Fanuc KAREL source: kd00006.KL

-- PROVISIONAL review KL for V770-1; original PC SHA256 f148d555a5ab890fe6bb85ac45592f87ae5cccf59ea5f73407380e3d84313837
-- Incomplete behavior may be omitted. Consult companion uncertainty JSON. Do not deploy.
PROGRAM KD00006
%NOLOCKGROUP
VAR
  I : INTEGER
  J : INTEGER
  B : BOOLEAN
  R : REAL
  S : STRING[80]
BEGIN
  -- UNRESOLVED_PC offsets 5-12; opcodes 9D,23
  -- UNRESOLVED_PC offsets 17-21; opcodes 7F
END KD00006
